Fanuc KAREL source: ka00040.KL

PROGRAM KA00040
%STACKSIZE=65535
%PRIORITY=65535
%NOLOCKGROUP
VAR
SRC : STRING[80]
DST : STRING[80]
BEGIN
SRC='A'
DST=SRC
END KA00040
